TYPE HmiCommand :
STRUCT
	sequence : UDINT;
	code : HmiCommandCode;
	manualTwist : Twist;
END_STRUCT
END_TYPE

(* stored: Version 1.1.0.1, ProductVersion 3.1.4026.12
   DUT HmiCommand: Id {78386c4a-ae37-569b-8ec1-a634655af4bc} *)
